(*
 * Simulacion_Trifasico_MPC_v8_M6_it10_opt_S71200.scl
 *
 * Base: Simulacion_Trifasico_MPC_v8_M6_it10_opt_OB100ms_DIAG.scl (PLC Coder 24.1,
 * variante f: Parametros_MPC_v8, M = 6, P = 200, tope de 10 iteraciones, Kr 18x3,
 * divisor desactivado, instrumentacion [DIAG] con RUNTIME).
 *
 * MODIFICADO para S7-1200 (memoria de trabajo). La ley de control no cambia:
 *  1. Kr, Hinv, Ac y Linv pasan a valores iniciales de la declaracion. Se
 *     elimina el bloque need_init, que las cargaba con 2144 asignaciones.
 *  2. rseq pasa de 600 a 3 elementos (solo se usan rseq[0..2]) y se elimina
 *     vseq (201 unos que no se usaban); v sigue valiendo 1.0.
 *  3. Se eliminan las copias QQ y RR: se leen directamente i0_qr.b_Q y i0_qr.b_R.
 *  4. Los arreglos de solo lectura pasan de VAR_INPUT (copia en cada llamada)
 *     a VAR_IN_OUT (referencia): qr.b_A, xgemv.b_A (x se elimina porque en qr
 *     siempre es el mismo arreglo que b_A), mpc_clipping.b_Mlim
 *     y b_Mrows, abs_g.x, b_abs.x, maximum2.x.
 *  5. Bloques con los nombres del proyecto (sufijo _MPC; MPC_3 -> MPC_Control).
 *  v2 (para bajar del 100 % en la CPU 1212C), resultados identicos:
 *  6. Ac separada en AcS (SINT, columnas 0..17, valores -1/0/1) y AcSlack (REAL,
 *     columna 18); cada producto suma la columna 18 al final, en el mismo orden.
 *  7. Se elimina U: en el lazo se usa -b_H (negacion exacta) y en el arranque
 *     en caliente se guarda en TL, que se recalcula antes de volver a leerse.
 *  8. qr factoriza en el sitio sobre RLinv (sin la copia c_A).
 *  9. RLinv, TL y b_D pasan a VAR_TEMP (4332 B de pila local; limite 6 KB).
 * 10. d_a pasa de INT a SINT (valores -1/0/1).
 *  LLAMAR DESDE UN OB CICLICO DE 100 ms. Requiere el DB global Diag_HIL.
 *
 * Model name                      : Simulacion_Trifasico_MPC_v6
 * Model version                   : 1.95
 * Model creator                   : Ivan
 * Model last modified by          : Ivan
 * Model last modified on          : Tue Sep 22 00:34:01 2026
 * Model sample time               : 0.01s
 * Subsystem name                  : Simulacion_Trifasico_MPC_v6/MPC_3
 * Subsystem sample time           : 0.01s
 * Simulink PLC Coder version      : 24.1 (R2024a) 19-Nov-2023
 * ST code generated on            : Tue Sep 22 02:35:18 2026
 *
 * Target IDE selection            : Siemens TIA Portal
 * Test Bench included             : No
 *
 * MODIFICADO (post-proceso), variante f: Parametros_MPC_v8 con M = 6 y tope de 10 iteraciones (P = 200):
 *  - Kr reducida de 18x600 a 18x3: 54 operaciones por ejecucion en lugar de 10800.
 *  - Contador en DB propio: PLCGlobalVarMPC.plc_ts_counter_MPC
 *  - Divisor desactivado: el MPC ejecuta en cada llamada.
 *    LLAMAR DESDE UN OB CICLICO DE 100 ms (100000 us).
 *
 * MODIFICADO: instrumentacion de tiempo con RUNTIME (lineas marcadas [DIAG]).
 *  - Mide el paso completo del MPC: estimador + QP + recorte.
 *  - Registra el estado del QP: iteraciones, llegadas al tope e infactibles.
 *  - Requiere el DB global Diag_HIL (Diag_HIL.scl) en el proyecto.
 *  - La ley de control no cambia.
 *
 *)
DATA_BLOCK PLCGlobalVarMPC
STRUCT
    plc_ts_counter_MPC: DINT;
END_STRUCT
BEGIN
END_DATA_BLOCK
FUNCTION_BLOCK abs_g_MPC
VAR_OUTPUT
    y: ARRAY [0..71] OF REAL;
END_VAR
VAR_IN_OUT
    x: ARRAY [0..71] OF REAL;   (* solo lectura *)
END_VAR
VAR
    k: DINT;
END_VAR
FOR k := 0 TO 71 DO
    y[k] := ABS(x[k]);
END_FOR;
END_FUNCTION_BLOCK
FUNCTION_BLOCK b_abs_MPC
VAR_OUTPUT
    y: ARRAY [0..18] OF REAL;
END_VAR
VAR_IN_OUT
    x: ARRAY [0..18] OF REAL;   (* solo lectura *)
END_VAR
VAR
    k: DINT;
END_VAR
FOR k := 0 TO 18 DO
    y[k] := ABS(x[k]);
END_FOR;
END_FUNCTION_BLOCK
FUNCTION_BLOCK maximum2_MPC
VAR_INPUT
    y: REAL;
END_VAR
VAR_OUTPUT
    ex: ARRAY [0..71] OF REAL;
END_VAR
VAR_IN_OUT
    x: ARRAY [0..71] OF REAL;   (* solo lectura *)
END_VAR
VAR
    k: DINT;
END_VAR
FOR k := 0 TO 71 DO
    ex[k] := MAX(IN1:=x[k], IN2:=y);
END_FOR;
END_FUNCTION_BLOCK
FUNCTION_BLOCK mpc_clipping_MPC
VAR_INPUT
    uk: ARRAY [0..2] OF REAL;
    uk1: ARRAY [0..2] OF REAL;
    b_uoff: ARRAY [0..2] OF REAL;
    b_ny: DINT;
    b_degrees: DINT;
END_VAR
VAR_OUTPUT
    uk_clipped: ARRAY [0..2] OF REAL;
END_VAR
VAR_IN_OUT
    b_Mlim: ARRAY [0..71] OF REAL;   (* solo lectura *)
    b_Mrows: ARRAY [0..71] OF DINT;  (* solo lectura *)
END_VAR
VAR
    nylim: DINT;
    umax: ARRAY [0..2] OF REAL;
    umin: ARRAY [0..2] OF REAL;
    dumin: ARRAY [0..2] OF REAL;
    dumax: ARRAY [0..2] OF REAL;
    iu: DINT;
    du: REAL;
    b_i: DINT;
    tmp: DINT;
    temp1: BOOL;
    temp2: BOOL;
    temp3: BOOL;
END_VAR
nylim := (400 * b_ny) + 1200;
uk_clipped[0] := uk[0];
umax[0] := 3.4028234663852886E+37;
umin[0] := -3.4028234663852886E+37;
dumin[0] := -3.4028234663852886E+37;
dumax[0] := 3.4028234663852886E+37;
uk_clipped[1] := uk[1];
umax[1] := 3.4028234663852886E+37;
umin[1] := -3.4028234663852886E+37;
dumin[1] := -3.4028234663852886E+37;
dumax[1] := 3.4028234663852886E+37;
uk_clipped[2] := uk[2];
umax[2] := 3.4028234663852886E+37;
umin[2] := -3.4028234663852886E+37;
dumin[2] := -3.4028234663852886E+37;
dumax[2] := 3.4028234663852886E+37;
FOR b_i := 0 TO 71 DO
    iu := b_Mrows[b_i];
    temp1 := FALSE;
    temp2 := FALSE;
    temp3 := FALSE;
    IF iu > (nylim - 1200) THEN
        IF iu <= (nylim - 1197) THEN
            iu := (iu - nylim) + 1199;
            umax[iu] := b_Mlim[b_i] + b_uoff[iu];
        ELSE
            temp3 := TRUE;
        END_IF;
    ELSE
        temp3 := TRUE;
    END_IF;
    IF temp3 THEN
        IF iu > (nylim - 600) THEN
            IF iu <= (nylim - 597) THEN
                iu := (iu - nylim) + 599;
                umin[iu] := ( -b_Mlim[b_i]) + b_uoff[iu];
            ELSE
                temp2 := TRUE;
            END_IF;
        ELSE
            temp2 := TRUE;
        END_IF;
    END_IF;
    IF temp2 THEN
        IF iu > nylim THEN
            IF iu <= (nylim + 3) THEN
                dumax[(iu - nylim) - 1] := b_Mlim[b_i];
            ELSE
                temp1 := TRUE;
            END_IF;
        ELSE
            temp1 := TRUE;
        END_IF;
    END_IF;
    IF temp1 THEN
        tmp := nylim + b_degrees;
        IF iu > (tmp - 1) THEN
            IF iu <= (tmp + 2) THEN
                dumin[(iu - nylim) - b_degrees] :=  -b_Mlim[b_i];
            END_IF;
        END_IF;
    END_IF;
END_FOR;
du := uk[0] - uk1[0];
IF du > dumax[0] THEN
    uk_clipped[0] := uk1[0] + dumax[0];
ELSIF du < dumin[0] THEN
    uk_clipped[0] := uk1[0] + dumin[0];
END_IF;
IF uk_clipped[0] > umax[0] THEN
    uk_clipped[0] := umax[0];
ELSIF uk_clipped[0] < umin[0] THEN
    uk_clipped[0] := umin[0];
END_IF;
du := uk[1] - uk1[1];
IF du > dumax[1] THEN
    uk_clipped[1] := uk1[1] + dumax[1];
ELSIF du < dumin[1] THEN
    uk_clipped[1] := uk1[1] + dumin[1];
END_IF;
IF uk_clipped[1] > umax[1] THEN
    uk_clipped[1] := umax[1];
ELSIF uk_clipped[1] < umin[1] THEN
    uk_clipped[1] := umin[1];
END_IF;
du := uk[2] - uk1[2];
IF du > dumax[2] THEN
    uk_clipped[2] := uk1[2] + dumax[2];
ELSIF du < dumin[2] THEN
    uk_clipped[2] := uk1[2] + dumin[2];
END_IF;
IF uk_clipped[2] > umax[2] THEN
    uk_clipped[2] := umax[2];
ELSIF uk_clipped[2] < umin[2] THEN
    uk_clipped[2] := umin[2];
END_IF;
END_FUNCTION_BLOCK
FUNCTION maximum_MPC: REAL
VAR_INPUT
    x: ARRAY [0..18] OF REAL;
END_VAR
VAR_TEMP
    k: DINT;
    x_0: REAL;
END_VAR
maximum_MPC := x[0];
FOR k := 0 TO 17 DO
    x_0 := x[k + 1];
    IF maximum_MPC < x_0 THEN
        maximum_MPC := x_0;
    END_IF;
END_FOR;
END_FUNCTION
FUNCTION_BLOCK DropConstraint_MPC
VAR_INPUT
    kDrop: DINT;
END_VAR
VAR_IN_OUT
    iA: ARRAY [0..71] OF BOOL;
    nA: DINT;
    iC: ARRAY [0..71] OF DINT;
END_VAR
VAR
    b_i: DINT;
END_VAR
IF kDrop > 0 THEN
    iA[iC[kDrop - 1] - 1] := FALSE;
    IF kDrop < nA THEN
        b_i := kDrop;
        WHILE b_i <= (nA - 1) DO
            iC[b_i - 1] := iC[b_i];
            b_i := b_i + 1;
        END_WHILE;
    END_IF;
    iC[nA - 1] := 0;
    nA := nA - 1;
END_IF;
END_FUNCTION_BLOCK
FUNCTION mtimes_MPC: REAL
VAR_INPUT
    b_A: ARRAY [0..18] OF REAL;
    B: ARRAY [0..18] OF REAL;
END_VAR
VAR_TEMP
    k: DINT;
END_VAR
mtimes_MPC := 0.0;
FOR k := 0 TO 18 DO
    mtimes_MPC := (b_A[k] * B[k]) + mtimes_MPC;
END_FOR;
END_FUNCTION
FUNCTION xnrm2_MPC: REAL
VAR_INPUT
    b_n: DINT;
    x: ARRAY [0..360] OF REAL;
    ix0: DINT;
END_VAR
VAR_TEMP
    b_scale: REAL;
    kend: DINT;
    absxk: REAL;
    t: REAL;
    k: DINT;
END_VAR
xnrm2_MPC := 0.0;
IF b_n >= 1 THEN
    IF b_n = 1 THEN
        xnrm2_MPC := ABS(x[ix0 - 1]);
    ELSE
        b_scale := 1.1754943508222875E-37;
        kend := (ix0 + b_n) - 1;
        k := ix0;
        WHILE k <= kend DO
            absxk := ABS(x[k - 1]);
            IF absxk > b_scale THEN
                t := b_scale / absxk;
                xnrm2_MPC := ((xnrm2_MPC * t) * t) + 1.0;
                b_scale := absxk;
            ELSE
                t := absxk / b_scale;
                xnrm2_MPC := (t * t) + xnrm2_MPC;
            END_IF;
            k := k + 1;
        END_WHILE;
        xnrm2_MPC := b_scale * SQRT(xnrm2_MPC);
    END_IF;
END_IF;
END_FUNCTION
FUNCTION_BLOCK xgerc_MPC
VAR_INPUT
    b_m: DINT;
    b_n: DINT;
    alpha1: REAL;
    ix0: DINT;
    y: ARRAY [0..18] OF REAL;
    ia0: DINT;
END_VAR
VAR_IN_OUT
    b_A: ARRAY [0..360] OF REAL;
END_VAR
VAR
    jA: DINT;
    jy: DINT;
    temp: REAL;
    ix: DINT;
    j: DINT;
    b_b: DINT;
    ijA: DINT;
END_VAR
IF alpha1 <> 0.0 THEN
    jA := ia0 - 1;
    jy := 0;
    j := 0;
    WHILE j <= (b_n - 1) DO
        IF y[jy] <> 0.0 THEN
            temp := y[jy] * alpha1;
            ix := ix0;
            ijA := jA;
            b_b := b_m + jA;
            WHILE (ijA + 1) <= b_b DO
                b_A[ijA] := (b_A[ix - 1] * temp) + b_A[ijA];
                ix := ix + 1;
                ijA := ijA + 1;
            END_WHILE;
        END_IF;
        jy := jy + 1;
        jA := jA + 19;
        j := j + 1;
    END_WHILE;
END_IF;
END_FUNCTION_BLOCK
FUNCTION_BLOCK xgemv_MPC
VAR_INPUT
    b_m: DINT;
    b_n: DINT;
    ia0: DINT;
    ix0: DINT;
END_VAR
VAR_IN_OUT
    y: ARRAY [0..18] OF REAL;
    b_A: ARRAY [0..360] OF REAL;   (* solo lectura, por referencia; hace tambien de x: en qr siempre x = b_A = c_A *)
END_VAR
VAR
    ix: DINT;
    b_c: REAL;
    b_iy: DINT;
    b_b: DINT;
    iac: DINT;
    b_d: DINT;
    ia: DINT;
END_VAR
IF (b_m <> 0) AND (b_n <> 0) THEN
    b_iy := 0;
    WHILE b_iy <= (b_n - 1) DO
        y[b_iy] := 0.0;
        b_iy := b_iy + 1;
    END_WHILE;
    b_iy := 0;
    b_b := ((b_n - 1) * 19) + ia0;
    iac := ia0;
    WHILE iac <= b_b DO
        ix := ix0;
        b_c := 0.0;
        b_d := (iac + b_m) - 1;
        ia := iac;
        WHILE ia <= b_d DO
            b_c := (b_A[ia - 1] * b_A[ix - 1]) + b_c;
            ix := ix + 1;
            ia := ia + 1;
        END_WHILE;
        y[b_iy] := y[b_iy] + b_c;
        b_iy := b_iy + 1;
        iac := iac + 19;
    END_WHILE;
END_IF;
END_FUNCTION_BLOCK
FUNCTION_BLOCK qr_MPC
VAR_OUTPUT
    b_Q: ARRAY [0..360] OF REAL;
    b_R: ARRAY [0..360] OF REAL;
END_VAR
VAR_IN_OUT
    b_A: ARRAY [0..360] OF REAL;   (* se factoriza en el sitio: el llamador no vuelve a leer RLinv sin ponerla a cero *)
END_VAR
VAR
    i0_xgemv: xgemv_MPC;
    i0_xgerc: xgerc_MPC;
    tau: ARRAY [0..18] OF REAL;
    itau: DINT;
    work: ARRAY [0..18] OF REAL;
    ii: DINT;
    atmp: REAL;
    beta1: REAL;
    knt: DINT;
    c_lastc: DINT;
    coltop: DINT;
    b_coltop: DINT;
    c_A_0: REAL;
    a: REAL;
    exitg1: DINT;
    exitg2: DINT;
    temp7: REAL;
END_VAR
FOR ii := 0 TO 18 DO
    tau[ii] := 0.0;
    work[ii] := 0.0;
END_FOR;
FOR itau := 0 TO 18 DO
    ii := (itau * 19) + itau;
    IF (itau + 1) < 19 THEN
        atmp := b_A[ii];
        tau[itau] := 0.0;
        beta1 := xnrm2_MPC(b_n := 18 - itau, x := b_A, ix0 := ii + 2);
        IF beta1 <> 0.0 THEN
            c_A_0 := b_A[ii];
            a := ABS(c_A_0);
            beta1 := ABS(beta1);
            IF a < beta1 THEN
                a := a / beta1;
                beta1 := SQRT((a * a) + 1.0) * beta1;
            ELSIF a > beta1 THEN
                beta1 := beta1 / a;
                beta1 := SQRT((beta1 * beta1) + 1.0) * a;
            ELSE
                beta1 := a * 1.4142135623730951;
            END_IF;
            IF c_A_0 >= 0.0 THEN
                beta1 :=  -beta1;
            END_IF;
            IF ABS(beta1) < 1.1754943508222875E-37 THEN
                knt := 0;
                REPEAT
                    exitg1 := 0;
                    knt := knt + 1;
                    c_lastc := (ii - itau) + 19;
                    b_coltop := ii + 1;
                    WHILE (b_coltop + 1) <= c_lastc DO
                        b_A[b_coltop] := 3.4028234663852886E+37 * b_A[b_coltop];
                        b_coltop := b_coltop + 1;
                    END_WHILE;
                    beta1 := beta1 * 3.4028234663852886E+37;
                    atmp := atmp * 3.4028234663852886E+37;
                    IF ABS(beta1) < 1.1754943508222875E-37 THEN
                        IF knt < 20 THEN
                            ;
                            ;
                        ELSE
                            exitg1 := 1;
                        END_IF;
                    ELSE
                        exitg1 := 1;
                    END_IF;
                UNTIL NOT(exitg1 = 0)
                END_REPEAT;
                a := ABS(atmp);
                temp7 := xnrm2_MPC(b_n := 18 - itau, x := b_A, ix0 := ii + 2);
                beta1 := ABS(temp7);
                IF a < beta1 THEN
                    a := a / beta1;
                    beta1 := SQRT((a * a) + 1.0) * beta1;
                ELSIF a > beta1 THEN
                    beta1 := beta1 / a;
                    beta1 := SQRT((beta1 * beta1) + 1.0) * a;
                ELSE
                    beta1 := a * 1.4142135623730951;
                END_IF;
                IF atmp >= 0.0 THEN
                    beta1 :=  -beta1;
                END_IF;
                tau[itau] := (beta1 - atmp) / beta1;
                atmp := 1.0 / (atmp - beta1);
                b_coltop := ii + 1;
                WHILE (b_coltop + 1) <= c_lastc DO
                    b_A[b_coltop] := atmp * b_A[b_coltop];
                    b_coltop := b_coltop + 1;
                END_WHILE;
                c_lastc := 0;
                WHILE c_lastc <= (knt - 1) DO
                    beta1 := beta1 * 1.1754943508222875E-37;
                    c_lastc := c_lastc + 1;
                END_WHILE;
                atmp := beta1;
            ELSE
                tau[itau] := (beta1 - c_A_0) / beta1;
                atmp := 1.0 / (c_A_0 - beta1);
                knt := (ii - itau) + 19;
                c_lastc := ii + 1;
                WHILE (c_lastc + 1) <= knt DO
                    b_A[c_lastc] := atmp * b_A[c_lastc];
                    c_lastc := c_lastc + 1;
                END_WHILE;
                atmp := beta1;
            END_IF;
        END_IF;
        b_A[ii] := 1.0;
        IF tau[itau] <> 0.0 THEN
            knt := 19 - itau;
            c_lastc := (ii - itau) + 18;
            REPEAT
                exitg1 := 0;
                IF knt > 0 THEN
                    IF b_A[c_lastc] = 0.0 THEN
                        knt := knt - 1;
                        c_lastc := c_lastc - 1;
                    ELSE
                        exitg1 := 1;
                    END_IF;
                ELSE
                    exitg1 := 1;
                END_IF;
            UNTIL NOT(exitg1 = 0)
            END_REPEAT;
            c_lastc := 18 - itau;
            REPEAT
                exitg2 := 0;
                IF c_lastc > 0 THEN
                    b_coltop := (((c_lastc - 1) * 19) + ii) + 19;
                    coltop := b_coltop;
                    REPEAT
                        exitg1 := 0;
                        IF (coltop + 1) <= (b_coltop + knt) THEN
                            IF b_A[coltop] <> 0.0 THEN
                                exitg1 := 1;
                            ELSE
                                coltop := coltop + 1;
                            END_IF;
                        ELSE
                            c_lastc := c_lastc - 1;
                            exitg1 := 2;
                        END_IF;
                    UNTIL NOT(exitg1 = 0)
                    END_REPEAT;
                    IF exitg1 = 1 THEN
                        exitg2 := 1;
                    END_IF;
                ELSE
                    exitg2 := 1;
                END_IF;
            UNTIL NOT(exitg2 = 0)
            END_REPEAT;
        ELSE
            knt := 0;
            c_lastc := 0;
        END_IF;
        IF knt > 0 THEN
            i0_xgemv(b_m := knt, b_n := c_lastc, b_A := b_A, ia0 := ii + 20, ix0 := ii + 1, y := work);
            i0_xgerc(b_m := knt, b_n := c_lastc, alpha1 :=  -tau[itau], ix0 := ii + 1, y := work, b_A := b_A, ia0 := ii + 20)
                ;
        END_IF;
        b_A[ii] := atmp;
    ELSE
        tau[18] := 0.0;
    END_IF;
END_FOR;
FOR itau := 0 TO 18 DO
    ii := 0;
    WHILE ii <= itau DO
        b_R[ii + (19 * itau)] := b_A[(19 * itau) + ii];
        ii := ii + 1;
    END_WHILE;
    ii := itau + 1;
    WHILE (ii + 1) < 20 DO
        b_R[ii + (19 * itau)] := 0.0;
        ii := ii + 1;
    END_WHILE;
    work[itau] := 0.0;
END_FOR;
FOR ii := 18 TO 0 BY -1 DO
    knt := ((ii * 19) + ii) + 20;
    IF (ii + 1) < 19 THEN
        b_A[knt - 20] := 1.0;
        IF tau[ii] <> 0.0 THEN
            c_lastc := 19 - ii;
            b_coltop := knt - ii;
            REPEAT
                exitg1 := 0;
                IF c_lastc > 0 THEN
                    IF b_A[b_coltop - 2] = 0.0 THEN
                        c_lastc := c_lastc - 1;
                        b_coltop := b_coltop - 1;
                    ELSE
                        exitg1 := 1;
                    END_IF;
                ELSE
                    exitg1 := 1;
                END_IF;
            UNTIL NOT(exitg1 = 0)
            END_REPEAT;
            b_coltop := 18 - ii;
            REPEAT
                exitg2 := 0;
                IF b_coltop > 0 THEN
                    coltop := ((b_coltop - 1) * 19) + knt;
                    itau := coltop;
                    REPEAT
                        exitg1 := 0;
                        IF itau <= ((coltop + c_lastc) - 1) THEN
                            IF b_A[itau - 1] <> 0.0 THEN
                                exitg1 := 1;
                            ELSE
                                itau := itau + 1;
                            END_IF;
                        ELSE
                            b_coltop := b_coltop - 1;
                            exitg1 := 2;
                        END_IF;
                    UNTIL NOT(exitg1 = 0)
                    END_REPEAT;
                    IF exitg1 = 1 THEN
                        exitg2 := 1;
                    END_IF;
                ELSE
                    exitg2 := 1;
                END_IF;
            UNTIL NOT(exitg2 = 0)
            END_REPEAT;
        ELSE
            c_lastc := 0;
            b_coltop := 0;
        END_IF;
        IF c_lastc > 0 THEN
            i0_xgemv(b_m := c_lastc, b_n := b_coltop, b_A := b_A, ia0 := knt, ix0 := knt - 19, y := work);
            i0_xgerc(b_m := c_lastc, b_n := b_coltop, alpha1 :=  -tau[ii], ix0 := knt - 19, y := work, b_A := b_A, ia0 := knt)
                ;
        END_IF;
        c_lastc := (knt - ii) - 1;
        b_coltop := knt - 19;
        WHILE (b_coltop + 1) <= c_lastc DO
            b_A[b_coltop] := ( -tau[ii]) * b_A[b_coltop];
            b_coltop := b_coltop + 1;
        END_WHILE;
    END_IF;
    b_A[knt - 20] := 1.0 - tau[ii];
    c_lastc := 0;
    WHILE c_lastc <= (ii - 1) DO
        b_A[(knt - c_lastc) - 21] := 0.0;
        c_lastc := c_lastc + 1;
    END_WHILE;
END_FOR;
FOR ii := 0 TO 360 DO
    b_Q[ii] := b_A[ii];
END_FOR;
END_FUNCTION_BLOCK
FUNCTION b_norm_MPC: REAL
VAR_INPUT
    x: ARRAY [0..18] OF REAL;
END_VAR
VAR_TEMP
    b_scale: REAL;
    absxk: REAL;
    t: REAL;
    k: DINT;
END_VAR
b_norm_MPC := 0.0;
b_scale := 1.1754943508222875E-37;
FOR k := 0 TO 18 DO
    absxk := ABS(x[k]);
    IF absxk > b_scale THEN
        t := b_scale / absxk;
        b_norm_MPC := ((b_norm_MPC * t) * t) + 1.0;
        b_scale := absxk;
    ELSE
        t := absxk / b_scale;
        b_norm_MPC := (t * t) + b_norm_MPC;
    END_IF;
END_FOR;
b_norm_MPC := b_scale * SQRT(b_norm_MPC);
END_FUNCTION
FUNCTION_BLOCK mpcblock_refmd_MPC
VAR_INPUT
    b_ref: ARRAY [0..2] OF REAL;
    b_yoff: ARRAY [0..2] OF REAL;
    b_RYscale: ARRAY [0..2] OF REAL;
END_VAR
VAR_OUTPUT
    rseq: ARRAY [0..2] OF REAL;   (* antes 0..599: solo se usan rseq[0..2] *)
    v: REAL;
END_VAR
VAR
    b_i: DINT;
    ref_0: REAL;
    ref_1: REAL;
    ref_2: REAL;
    b_RYscale_0: REAL;
    b_RYscale_1: REAL;
    b_RYscale_2: REAL;
    b_yoff_0: REAL;
    b_yoff_1: REAL;
    b_yoff_2: REAL;
END_VAR
ref_0 := b_ref[0];
ref_1 := b_ref[1];
ref_2 := b_ref[2];
b_RYscale_0 := b_RYscale[0];
b_RYscale_1 := b_RYscale[1];
b_RYscale_2 := b_RYscale[2];
b_yoff_0 := b_yoff[0];
b_yoff_1 := b_yoff[1];
b_yoff_2 := b_yoff[2];
FOR b_i := 0 TO 0 DO    (* solo rseq[0..2] se usa *)
    rseq[b_i * 3] := (ref_0 * b_RYscale_0) - b_yoff_0;
    rseq[(b_i * 3) + 1] := (ref_1 * b_RYscale_1) - b_yoff_1;
    rseq[(b_i * 3) + 2] := (ref_2 * b_RYscale_2) - b_yoff_2;
END_FOR;
v := 1.0;
END_FUNCTION_BLOCK
FUNCTION rt_floord_MPC: REAL
VAR_INPUT
    u: REAL;
END_VAR
rt_floord_MPC := DINT_TO_REAL(TRUNC(u));
IF u = rt_floord_MPC THEN
    rt_floord_MPC := u;
ELSIF u < 0.0 THEN
    rt_floord_MPC := rt_floord_MPC - 1.0;
END_IF;
END_FUNCTION
FUNCTION_BLOCK MPC_Control
VAR_INPUT
    ssMethodType: INT;
    moorx: ARRAY [0..2] OF REAL;
    b_ref: ARRAY [0..2] OF REAL;
END_VAR
VAR_OUTPUT
    mv: ARRAY [0..2] OF REAL;
END_VAR
VAR
    Memory_PreviousInput: ARRAY [0..71] OF BOOL;
    last_x_PreviousInput: ARRAY [0..6] OF REAL;
    last_mv_DSTATE: ARRAY [0..2] OF REAL;
    MathFunction: ARRAY [0..2] OF REAL;
    MathFunction1: ARRAY [0..2] OF REAL;
    MathFunction2: ARRAY [0..2] OF REAL;
    c_last_x_InitialCond: ARRAY [0..6] OF REAL := [0.47374550049727165,0.8,0.72,255106.009,0.0,0.0,0.0];
    MPC_3_b_myoff: ARRAY [0..2] OF REAL := [0.8,0.72,3.7];
    MPC_3_b_RYscale: ARRAY [0..2] OF REAL := [1.0,1.0,0.1];
    MPC_3_b_xoff: ARRAY [0..6] OF REAL := [0.47374550049727165,0.8,0.72,255106.009,0.0,0.0,0.0];
    b_a: ARRAY [0..20] OF REAL := [0.0,0.0,0.0,1.0,0.0,0.0,0.0,1.0,0.0,0.0,0.0,1.4503774389728313E-5,0.0,0.0,0.0,0.0,0.0,0.0,0.0,
        0.0,0.0];
    MPC_3_c_a: ARRAY [0..20] OF REAL := [-0.0772292027423523,0.12077646327456022,0.0038948707411090538,1352.9330397447068,
        3.4881337436777948,-1.3447885799979777,-1.1731438171327024,0.269035613232814,0.0038948707411099914,0.09786695730401461,
        348.05070726193321,0.11111867957141662,2.7949959088743932,-2.8155753844244291,0.059593437249509731,0.01962263557286395,
        0.0050480489343075492,14331.413461436903,1.6106730948140586,2.3311020292522353,2.408935193579286];
    d_a: ARRAY [0..215] OF SINT := [-1,0,0,-1,0,0,-1,0,0,-1,0,0,-1,0,0,-1,0,0,1,0,0,1,0,0,1,0,0,1,0,0,1,0,0,1,0,0,0,0,0,0,0,0,0,0,0,
        0,0,0,0,0,0,0,0,0,0,0,0,0,0,0,0,0,0,0,0,0,0,0,0,0,0,0,0,-1,0,0,-1,0,0,-1,0,0,-1,0,0,-1,0,0,-1,0,0,1,0,0,1,0,0,1,0,0,
        1,0,0,1,0,0,1,0,0,0,0,0,0,0,0,0,0,0,0,0,0,0,0,0,0,0,0,0,0,0,0,0,0,0,0,0,0,0,0,0,0,0,0,0,0,0,-1,0,0,-1,0,0,-1,0,0,-1,
        0,0,-1,0,0,-1,0,0,1,0,0,1,0,0,1,0,0,1,0,0,1,0,0,1,0,0,0,0,0,0,0,0,0,0,0,0,0,0,0,0,0,0,0,0,0,0,0,0,0,0,0,0,0,0,0,0,0,
        0,0,0];
    MPC_3_b_Mlim: ARRAY [0..71] OF REAL := [0.333871875208127,0.752014397384409,0.515635973890735,0.333871875208127,
        0.752014397384409,0.515635973890735,0.333871875208127,0.752014397384409,0.515635973890735,0.333871875208127,0.752014397384409,
        0.515635973890735,0.333871875208127,0.752014397384409,0.515635973890735,0.333871875208127,0.752014397384409,0.515635973890735,
        0.636128124791873,0.21798560261559102,0.45436402610926496,0.636128124791873,0.21798560261559102,0.45436402610926496,
        0.636128124791873,0.21798560261559102,0.45436402610926496,0.636128124791873,0.21798560261559102,0.45436402610926496,
        0.636128124791873,0.21798560261559102,0.45436402610926496,0.636128124791873,0.21798560261559102,0.45436402610926496,0.035,0.015,
        0.03,0.035,0.015,0.03,0.035,0.015,0.03,0.035,0.015,0.03,0.035,0.015,0.03,0.035,0.015,0.03,0.035,0.015,0.03,0.035,0.015,
        0.03,0.035,0.015,0.03,0.035,0.015,0.03,0.035,0.015,0.03,0.035,0.015,0.03];
    MPC_3_b_Kx: ARRAY [0..125] OF REAL := [-7716.2321024491939,-10901.008671532656,-4264.9443651421188,0.001588040838629834,
        -2543.7442519006345,-1928.3474040587275,19.549174933816971,-44534.108859815329,-44494.776516572136,-26655.405567238093,
        0.0095121063518449449,-8398.6455416316712,-10368.267059564856,158.86185382546796,877.70571831208667,990.07022975809957,
        474.28108255756024,-0.0035701887162486057,96.5496604150103,99.981804413078876,-126.88330315000997,-7621.9188571763643,
        -10775.120625744157,-4206.5654308225376,0.0015700336455973293,-2519.1535379237243,-1907.0052261791157,19.280661326360363,
        -44188.119848216615,-44149.311125111242,-26390.969999054745,0.0094459267062587185,-8342.2703225681144,-10298.597291206755,
        157.85188650166057,864.95022738088733,975.66168439016542,466.81791298662728,-0.0035336819710021609,94.4868041100247,
        97.85316386731445,-125.93879584019494,-7528.1481322542822,-10649.931335099882,-4148.6767278274638,0.0015521046865827432,
        -2494.6400124657093,-1885.7587961853874,19.013959064141872,-43842.116288935795,-43803.826542255309,-26127.843886728973,
        0.0093796925467878947,-8285.8873550992248,-10228.919297363989,156.8419334382582,852.3095979437818,961.384106890396,459.43616436780036,
        -0.003497369852713806,92.447632839384539,95.74911914998566,-124.99418234183436,-7434.9230075303494,-10525.443894660129,
        -4091.2769580451954,0.0015342547665065048,-2470.2045128943837,-1864.6086925692725,18.749068146716176,-43496.122480806749,
        -43458.347088410825,-25866.027371158609,0.0093134067140901722,-8229.4967444644935,-10159.23320514503,155.83198146211291,
        839.78359704931961,947.23718912342133,452.13534732790527,-0.0034612522993006938,90.432068275420264,93.669582511506164,
        -124.04951211934259,-7342.2465048437853,-10401.661341488485,-4034.3648155478659,0.0015164846849855819,-2445.8478788030538,
        -1843.5554965261258,18.485988665509439,-43150.162591337648,-43112.896952629555,-25605.520593125708,0.0092470720701684772,
        -8173.0986508239621,-10089.539209226115,154.82201815145478,827.37198501561852,933.22061617028339,444.91497290855955,
        -0.0034253292477243787,88.440031602080353,91.614465843510473,-123.10483463065196,-7250.1215881048793,-10278.586654731167,
        -3977.9389865477651,0.00149879523623798,-2421.5709518529893,-1822.5997917608677,18.224720801734843,-42804.2606574284,
        -42767.500193326021,-25346.323693295184,0.0091806914982297729,-8116.6932889508143,-10019.83757147498,153.81203184149854,
        815.07451548496078,919.33406638300414,437.7745525706747,-0.0033896006339887937,86.47144350229388,89.5836806634611,
        -122.16019932703135];
    MPC_3_b_Ku1: ARRAY [0..53] OF REAL := [532.9519035819452,1758.7630386838541,-20.218495148255496,1758.7630386838541,
        9920.4082612993716,-164.30092992093171,-20.218495148255496,-164.30092992093171,131.49311423922407,527.80102628666316,
        1737.934860701725,-19.940788232849528,1746.9574860985949,9846.5918503106168,-163.25638356511735,-19.786511752201875,
        -161.71101778484783,130.514941055735,522.666313063715,1717.21838942958,-19.664954679108821,1735.1503109173054,9772.77075083077,
        -162.21185195795246,-19.359488246736596,-159.14605147852319,129.53665804804106,517.54793926655793,1696.6142696551719,
        -19.390994486572826,1723.3415351782228,9698.9487212665517,-161.16732147527,-18.93740822923742,-156.60596908182839,128.55831637410802,
        512.44608071469349,1676.1231380934234,-19.118907749797927,1711.5311924205112,9625.129520129678,-160.12277927000616,
        -18.520255194809877,-154.09070753671722,127.57996718519767,507.36091366067569,1655.7456233405144,-18.848694656201634,
        1699.7193276198914,9551.3169060341625,-159.07821327799945,-18.108012533640888,-151.60020265098143,126.60166162568011];
    MPC_3_b_Kr: ARRAY [0..53] OF REAL := [3186.8373350513389,4275.3677914960599,51.13509990647421,-32.452540397628589,26714.198696645544,72.918687149547608,
        -112.44555961175674,-475.25673471668864,252.72878690712173,3155.2425613858004,4216.8654170260106,50.638144210838703,
        -31.975100691061328,26449.325655557303,72.210143687081711,-110.79080635121332,-467.77820186026861,250.27164490947899,
        3123.8040857581582,4158.8539359264387,50.143499486122451,-31.502311016836352,26185.762042540995,71.504893608304656,
        -109.15217877028672,-460.38123779321489,247.82594499281888,3092.5219240585361,4101.3320539069082,49.651167400702548,
        -31.034149716397167,25923.508020768073,70.802939302930895,-107.52960162200367,-453.06535277614643,245.39169524300604,
        3061.396092190324,4044.2984688129827,49.161149624113243,-30.57059511536292,25662.563753294817,70.104283162373875,
        -105.92299960583885,-445.83005747772961,242.96890375165114,3030.4266060701984,3987.7518705822636,48.673447827046601,
        -30.111625523516803,25402.929403061011,69.408927579747242,-104.33229736767574,-438.67486297920362,240.55757861611488];   (* Kr reducida 18x3 *)
    MPC_3_b_Hinv: ARRAY [0..360] OF REAL := [0.1702344980572631,-0.000316051953237396,-0.0001214533827540456,-0.036345548841276047,-0.00022994447282000675,
        -7.8535204077971989E-5,-0.035434727013087031,-0.00014382977097906262,-3.4945956300716842E-5,-0.034542309014010772,
        -5.7720706811642746E-5,8.813456011776322E-6,-0.03366968301464044,2.8361008307101794E-5,5.2380161360600679E-5,
        -0.032817675154182616,0.00011438593593406882,9.552481608298865E-5,0.0,-0.000316051953237396,0.010547207252793461,
        2.1132487152157335E-5,-0.0001808791608454948,-0.0023314158969080174,1.0330320315621911E-5,-4.9534035220164727E-5,
        -0.0022413766833578007,1.2191170747377299E-7,7.8036147649309862E-5,-0.0021522792952646508,-9.54953740575078E-6,
        0.00020190252942289518,-0.0020644122541486152,-1.8729858790232883E-5,0.0003221473455128597,-0.0019779594821308214,
        -2.7454115420488076E-5,0.0,-0.0001214533827540456,2.1132487152157335E-5,0.30304411821884769,-6.514990994147179E-5,
        2.1728353827661485E-5,-0.064405415788092474,-8.97885060327611E-6,2.2273463510311548E-5,-0.062989706993492336,
        4.65603793551569E-5,2.2723267969727878E-5,-0.061614542822731315,0.00010110834451599296,2.3046591530932414E-5,
        -0.060282635561179215,0.00015444098334013595,2.322473034505095E-5,-0.058995530723217567,0.0,-0.036345548841276047,
        -0.0001808791608454948,-6.514990994147179E-5,0.17176291685304779,-0.00013612744730930092,-4.4560767159202152E-5,
        -0.0350971665966896,-9.13556293645426E-5,-2.2988766629637194E-5,-0.034463114486899891,-4.65576358502461E-5,
        -9.4991020623304764E-7,-0.033843716347050953,-1.7392388529733022E-6,2.1176229123452892E-5,-0.033239892629933931,
        4.3085064069324768E-5,4.3143636253156359E-5,0.0,-0.00022994447282000675,-0.0023314158969080174,2.1728353827661485E-5,
        -0.00013612744730930092,0.010698246530635966,1.2340538427932472E-5,-4.4760194642908621E-5,-0.0022102015392433554,
        3.4084100679808667E-6,4.4173612422238355E-5,-0.00214976861316072,-5.120830508461208E-6,0.00013070925637258645,
        -0.0020899593246978244,-1.3289405671251868E-5,0.00021489433364024608,-0.0020309671075964997,-2.1128873179308238E-5,
        0.0,-7.8535204077971989E-5,1.0330320315621911E-5,-0.064405415788092474,-4.4560767159202152E-5,1.2340538427932472E-5,
        0.3054148208775625,-1.015071319787011E-5,1.4368446176665112E-5,-0.062417276373171432,2.4179024444158472E-5,
        1.636636500723434E-5,-0.061380921474166857,5.8051555293553663E-5,1.8300251292219083E-5,-0.0603809302382588,
        9.1225498596546247E-5,2.0148793762691288E-5,-0.0594190724227041,0.0,-0.035434727013087031,-4.9534035220164727E-5,
        -8.97885060327611E-6,-0.0350971665966896,-4.4760194642908621E-5,-1.015071319787011E-5,0.17273845134311319,
        -3.9976889795088581E-5,-1.0826124612172019E-5,-0.034391366089294419,-3.5166046909618539E-5,-1.0727884762180431E-5,
        -0.0340234548514619,-3.0316948364924829E-5,-1.0252653775071641E-5,-0.033666135978688227,-2.5428615172775216E-5,
        -9.6634672683266118E-6,0.0,-0.00014382977097906262,-0.0022413766833578007,2.2273463510311548E-5,-9.13556293645426E-5,
        -0.0022102015392433554,1.4368446176665112E-5,-3.9976889795088581E-5,0.010790253977071384,6.7106504165377462E-6,
        1.0310200452023578E-5,-0.002147190141859824,-6.7830888060647946E-7,5.9505058354541645E-5,-0.0021154443640503916,
        -7.8370437343924534E-6,0.00010762063469870516,-0.0020839183592772296,-1.4793606326937087E-5,0.0,
        -3.4945956300716842E-5,1.2191170747377299E-7,-0.062989706993492336,-2.2988766629637194E-5,3.4084100679808667E-6,
        -0.062417276373171432,-1.0826124612172019E-5,6.7106504165377462E-6,0.30702802540700186,1.820897001919164E-6,
        1.005184108764361E-5,-0.061176025329871223,1.4557473121748288E-5,1.3395015801887418E-5,-0.060507679924504308,
        2.7124492071147717E-5,1.6716205009836463E-5,-0.059870813633310996,0.0,-0.034542309014010772,7.8036147649309862E-5,
        4.65603793551569E-5,-0.034463114486899891,4.4173612422238355E-5,2.4179024444158472E-5,-0.034391366089294419,
        1.0310200452023578E-5,1.820897001919164E-6,0.17318140332130527,-2.3547509119607678E-5,-2.0255119613621428E-5,
        -0.03420782335043554,-5.7379181065111574E-5,-4.1654408632959635E-5,-0.034095412692558565,-9.1167816691611789E-5,
        -6.2657366574418234E-5,0.0,-5.7720706811642746E-5,-0.0021522792952646508,2.2723267969727878E-5,-4.65576358502461E-5,
        -0.00214976861316072,1.636636500723434E-5,-3.5166046909618539E-5,-0.002147190141859824,1.005184108764361E-5,
        -2.3547509119607678E-5,0.010824871877124352,3.8016754445631412E-6,-1.1714654534696886E-5,-0.0021406660168113629,
        -2.3487140810286621E-6,3.1080884145891323E-7,-0.0021366194369659398,-8.4238697344242429E-6,0.0,8.813456011776322E-6,
        -9.54953740575078E-6,-0.061614542822731315,-9.4991020623304764E-7,-5.120830508461208E-6,-0.061380921474166857,
        -1.0727884762180431E-5,-6.7830888060647946E-7,-0.061176025329871223,-2.0255119613621428E-5,3.8016754445631412E-6,
        0.30790449828673894,-2.9132918265929341E-5,8.3532488641258142E-6,-0.060660620175687734,-3.7638527243085177E-5,
        1.2949735033266653E-5,-0.060348692971084965,0.0,-0.03366968301464044,0.00020190252942289518,0.00010110834451599296,
        -0.033843716347050953,0.00013070925637258645,5.8051555293553663E-5,-0.0340234548514619,5.9505058354541645E-5,
        1.4557473121748288E-5,-0.03420782335043554,-1.1714654534696886E-5,-2.9132918265929341E-5,0.17311211771562424,
        -8.2943372514784056E-5,-7.26451760390996E-5,-0.034526178406331057,-0.00015415495715396418,-0.00011546864934107219,0.0,
        2.8361008307101794E-5,-0.0020644122541486152,2.3046591530932414E-5,-1.7392388529733022E-6,-0.0020899593246978244,
        1.8300251292219083E-5,-3.0316948364924829E-5,-0.0021154443640503916,1.3395015801887418E-5,-5.7379181065111574E-5,
        -0.0021406660168113629,8.3532488641258142E-6,-8.2943372514784056E-5,0.010803886559746703,3.2103542526533054E-6,
        -0.00010704208143625654,-0.0021887753347569921,-1.9842771425297006E-6,0.0,5.2380161360600679E-5,
        -1.8729858790232883E-5,-0.060282635561179215,2.1176229123452892E-5,-1.3289405671251868E-5,-0.0603809302382588,
        -1.0252653775071641E-5,-7.8370437343924534E-6,-0.060507679924504308,-4.1654408632959635E-5,-2.3487140810286621E-6,
        -0.060660620175687734,-7.26451760390996E-5,3.2103542526533054E-6,0.308065547905881,-0.00010270880655031663,
        8.8847998121922669E-6,-0.0608495071191091,0.0,-0.032817675154182616,0.0003221473455128597,0.00015444098334013595,
        -0.033239892629933931,0.00021489433364024608,9.1225498596546247E-5,-0.033666135978688227,0.00010762063469870516,
        2.7124492071147717E-5,-0.034095412692558565,3.1080884145891323E-7,-3.7638527243085177E-5,-0.034526178406331057,
        -0.00010704208143625654,-0.00010270880655031663,0.17255097784265849,-0.00021442620951791223,-0.00016759605920454502,
        0.0,0.00011438593593406882,-0.0019779594821308214,2.322473034505095E-5,4.3085064069324768E-5,-0.0020309671075964997,
        2.0148793762691288E-5,-2.5428615172775216E-5,-0.0020839183592772296,1.6716205009836463E-5,-9.1167816691611789E-5,
        -0.0021366194369659398,1.2949735033266653E-5,-0.00015415495715396418,-0.0021887753347569921,8.8847998121922669E-6,
        -0.00021442620951791223,0.010729219465504205,4.5706825441767981E-6,0.0,9.552481608298865E-5,-2.7454115420488076E-5,
        -0.058995530723217567,4.3143636253156359E-5,-2.1128873179308238E-5,-0.0594190724227041,-9.6634672683266118E-6,
        -1.4793606326937087E-5,-0.059870813633310996,-6.2657366574418234E-5,-8.4238697344242429E-6,-0.060348692971084965,
        -0.00011546864934107219,-1.9842771425297006E-6,-0.0608495071191091,-0.00016759605920454502,4.5706825441767981E-6,
        0.30753298042695221,0.0,0.0,0.0,0.0,0.0,0.0,0.0,0.0,0.0,0.0,0.0,0.0,0.0,0.0,0.0,0.0,0.0,0.0,0.0,
        9.9999999999999974E-6];
    (* Ac (72 x 19, por columnas) separada: columnas 0..17 solo valen -1, 0 o 1 *)
    AcS: ARRAY [0..1295] OF SINT := [-1,0,0,-1,0,0,-1,0,0,-1,0,0,-1,0,0,-1,0,0,1,0,0,1,0,0,1,0,0,1,0,0,1,0,0,1,0,0,-1,0,0,0,0,0,0,0,0,0,0,0,0,0,0,0,0,0,1,
        0,0,0,0,0,0,0,0,0,0,0,0,0,0,0,0,0,0,-1,0,0,-1,0,0,-1,0,0,-1,0,0,-1,0,0,-1,0,0,1,0,0,1,0,0,1,0,0,1,0,0,1,0,0,1,0,0,-1,
        0,0,0,0,0,0,0,0,0,0,0,0,0,0,0,0,0,1,0,0,0,0,0,0,0,0,0,0,0,0,0,0,0,0,0,0,-1,0,0,-1,0,0,-1,0,0,-1,0,0,-1,0,0,-1,0,0,1,0,
        0,1,0,0,1,0,0,1,0,0,1,0,0,1,0,0,-1,0,0,0,0,0,0,0,0,0,0,0,0,0,0,0,0,0,1,0,0,0,0,0,0,0,0,0,0,0,0,0,0,0,0,0,0,-1,0,0,-1,
        0,0,-1,0,0,-1,0,0,-1,0,0,0,0,0,1,0,0,1,0,0,1,0,0,1,0,0,1,0,0,0,0,0,-1,0,0,0,0,0,0,0,0,0,0,0,0,0,0,0,0,0,1,0,0,0,0,0,0,
        0,0,0,0,0,0,0,0,0,0,0,0,-1,0,0,-1,0,0,-1,0,0,-1,0,0,-1,0,0,0,0,0,1,0,0,1,0,0,1,0,0,1,0,0,1,0,0,0,0,0,-1,0,0,0,0,0,0,0,
        0,0,0,0,0,0,0,0,0,0,1,0,0,0,0,0,0,0,0,0,0,0,0,0,0,0,0,0,0,-1,0,0,-1,0,0,-1,0,0,-1,0,0,-1,0,0,0,0,0,1,0,0,1,0,0,1,0,0,
        1,0,0,1,0,0,0,0,0,-1,0,0,0,0,0,0,0,0,0,0,0,0,0,0,0,0,0,1,0,0,0,0,0,0,0,0,0,0,0,0,0,0,0,0,0,0,-1,0,0,-1,0,0,-1,0,0,-1,
        0,0,0,0,0,0,0,0,1,0,0,1,0,0,1,0,0,1,0,0,0,0,0,0,0,0,-1,0,0,0,0,0,0,0,0,0,0,0,0,0,0,0,0,0,1,0,0,0,0,0,0,0,0,0,0,0,0,0,
        0,0,0,0,0,-1,0,0,-1,0,0,-1,0,0,-1,0,0,0,0,0,0,0,0,1,0,0,1,0,0,1,0,0,1,0,0,0,0,0,0,0,0,-1,0,0,0,0,0,0,0,0,0,0,0,0,0,0,
        0,0,0,1,0,0,0,0,0,0,0,0,0,0,0,0,0,0,0,0,0,0,-1,0,0,-1,0,0,-1,0,0,-1,0,0,0,0,0,0,0,0,1,0,0,1,0,0,1,0,0,1,0,0,0,0,0,0,0,
        0,-1,0,0,0,0,0,0,0,0,0,0,0,0,0,0,0,0,0,1,0,0,0,0,0,0,0,0,0,0,0,0,0,0,0,0,0,0,-1,0,0,-1,0,0,-1,0,0,0,0,0,0,0,0,0,0,0,1,
        0,0,1,0,0,1,0,0,0,0,0,0,0,0,0,0,0,-1,0,0,0,0,0,0,0,0,0,0,0,0,0,0,0,0,0,1,0,0,0,0,0,0,0,0,0,0,0,0,0,0,0,0,0,0,-1,0,0,
        -1,0,0,-1,0,0,0,0,0,0,0,0,0,0,0,1,0,0,1,0,0,1,0,0,0,0,0,0,0,0,0,0,0,-1,0,0,0,0,0,0,0,0,0,0,0,0,0,0,0,0,0,1,0,0,0,0,0,
        0,0,0,0,0,0,0,0,0,0,0,0,0,-1,0,0,-1,0,0,-1,0,0,0,0,0,0,0,0,0,0,0,1,0,0,1,0,0,1,0,0,0,0,0,0,0,0,0,0,0,-1,0,0,0,0,0,0,0,
        0,0,0,0,0,0,0,0,0,0,1,0,0,0,0,0,0,0,0,0,0,0,0,0,0,0,0,0,0,-1,0,0,-1,0,0,0,0,0,0,0,0,0,0,0,0,0,0,1,0,0,1,0,0,0,0,0,0,0,
        0,0,0,0,0,0,0,-1,0,0,0,0,0,0,0,0,0,0,0,0,0,0,0,0,0,1,0,0,0,0,0,0,0,0,0,0,0,0,0,0,0,0,0,0,-1,0,0,-1,0,0,0,0,0,0,0,0,0,
        0,0,0,0,0,1,0,0,1,0,0,0,0,0,0,0,0,0,0,0,0,0,0,-1,0,0,0,0,0,0,0,0,0,0,0,0,0,0,0,0,0,1,0,0,0,0,0,0,0,0,0,0,0,0,0,0,0,0,
        0,0,-1,0,0,-1,0,0,0,0,0,0,0,0,0,0,0,0,0,0,1,0,0,1,0,0,0,0,0,0,0,0,0,0,0,0,0,0,-1,0,0,0,0,0,0,0,0,0,0,0,0,0,0,0,0,0,1,
        0,0,0,0,0,0,0,0,0,0,0,0,0,0,0,0,0,0,-1,0,0,0,0,0,0,0,0,0,0,0,0,0,0,0,0,0,1,0,0,0,0,0,0,0,0,0,0,0,0,0,0,0,0,0,-1,0,0,0,
        0,0,0,0,0,0,0,0,0,0,0,0,0,0,1,0,0,0,0,0,0,0,0,0,0,0,0,0,0,0,0,0,0,-1,0,0,0,0,0,0,0,0,0,0,0,0,0,0,0,0,0,1,0,0,0,0,0,0,
        0,0,0,0,0,0,0,0,0,0,0,-1,0,0,0,0,0,0,0,0,0,0,0,0,0,0,0,0,0,1,0,0,0,0,0,0,0,0,0,0,0,0,0,0,0,0,0,0,-1,0,0,0,0,0,0,0,0,0,
        0,0,0,0,0,0,0,0,1,0,0,0,0,0,0,0,0,0,0,0,0,0,0,0,0,0,-1,0,0,0,0,0,0,0,0,0,0,0,0,0,0,0,0,0,1];
    AcSlack: ARRAY [0..71] OF REAL := [0.1,0.1,0.1,0.1,0.1,0.1,0.1,0.1,0.1,0.1,0.1,0.1,0.1,0.1,0.1,0.1,0.1,0.1,0.1,0.1,0.1,0.1,0.1,0.1,0.1,0.1,0.1,0.1,0.1,
        0.1,0.1,0.1,0.1,0.1,0.1,0.1,0.0,0.0,0.0,0.0,0.0,0.0,0.0,0.0,0.0,0.0,0.0,0.0,0.0,0.0,0.0,0.0,0.0,0.0,0.0,0.0,0.0,0.0,
        0.0,0.0,0.0,0.0,0.0,0.0,0.0,0.0,0.0,0.0,0.0,0.0,0.0,0.0];   (* columna 18: holgura *)
    MPC_3_b_uoff: ARRAY [0..2] OF REAL := [0.656128124791873,0.237985602615591,0.474364026109265];
    MPC_3_b_Mrows: ARRAY [0..71] OF DINT := [1201,1202,1203,1204,1205,1206,1207,1208,1209,1210,1211,1212,1213,1214,1215,1216,1217,
        1218,1801,1802,1803,1804,1805,1806,1807,1808,1809,1810,1811,1812,1813,1814,1815,1816,1817,1818,2401,2402,2403,2404,
        2405,2406,2407,2408,2409,2410,2411,2412,2413,2414,2415,2416,2417,2418,2419,2420,2421,2422,2423,2424,2425,2426,2427,
        2428,2429,2430,2431,2432,2433,2434,2435,2436];
    MPC_3_b_Linv: ARRAY [0..360] OF REAL := [0.043122239395521268,-0.05019306519247696,-0.0033206696132972837,-0.31577942830214772,-0.0031471197006212965,
        -0.00020705051348992359,-0.18308150772189805,-0.0014696017526715675,-7.5450474722372636E-5,-0.12889586192277314,
        -0.00059021717051271558,3.8407404253082784E-6,-0.09869296350827321,0.0002261820630442589,8.3395085100205E-5,
        -0.078999376861682777,0.0011042900946144102,0.00017225441484848154,0.0,0.0,0.015347363356332721,0.0020190838633724136,
        -0.00091102072052030891,-0.07901358568341027,6.7218935720810737E-5,-9.1246872819404E-6,-0.045684177963437142,
        -3.9801617956080181E-6,0.00027433939577582988,-0.031987683695103353,-2.7972250421381947E-5,0.00047973300959174817,
        -0.024247405963223941,-4.0683462098209086E-5,0.0006803357457738446,-0.01909559690027262,-4.9506429646829944E-5,0.0,
        0.0,0.0,0.087312641366686636,-0.00043386070373357613,0.001238779140346204,-0.42107641020149239,-6.1807887311560788E-5,
        0.00051363050814862469,-0.24423350048424408,7.3761326011918756E-5,0.00035445285917561705,-0.17220651542065402,
        0.00018273894349911022,0.00028329895418285477,-0.13225134353194426,0.00029556006650442523,0.00023268095887176668,
        -0.10638325243751168,0.0,0.0,0.0,0.0,0.32476352152728083,-0.0022032755395640763,-0.00021807552222073261,
        -0.1826323676701698,-0.0012233193115584247,-0.00011214950035355466,-0.12907314160690159,-0.00073675201931614072,
        -5.3944104655688172E-5,-0.0993319703512495,-0.00021614122189525552,6.5016994885151178E-6,-0.080019318890644078,
        0.00041594529543757932,7.77984415145777E-5,0.0,0.0,0.0,0.0,0.0,0.081196332633548682,9.4178408876197282E-5,
        -0.00018552342484247817,-0.045616373263034124,1.3382645905252523E-5,7.3265273574636073E-5,-0.032161700136474826,
        -1.4106521576734893E-5,0.00024883046634005361,-0.024605618012537182,-2.8451514186729147E-5,0.00041959371575441944,
        -0.019607343607742585,-3.810048357222283E-5,0.0,0.0,0.0,0.0,0.0,0.0,0.43311489522212737,-0.00017825206901915394,
        0.00037846148477057873,-0.24327007517811419,-5.0314671809548014E-5,0.00026963086606063725,-0.17200596953896155,
        4.5079990938181534E-5,0.0002299643325305634,-0.13258611861207259,0.00014267226685941574,0.00020304604787921979,
        -0.10714700086017916,0.0,0.0,0.0,0.0,0.0,0.0,0.0,0.37344065756375838,-0.00097294854471077308,-0.00014891231274351814,
        -0.12927510944801096,-0.00087014142142283494,-0.00011208292497242445,-0.099986751616224556,-0.00063795107819119646,
        -7.0970441026343978E-5,-0.081048819235342642,-0.00024549134958053907,-1.7425575551665338E-5,0.0,0.0,0.0,0.0,0.0,0.0,
        0.0,0.0,0.093363604583182686,3.0799370827412689E-5,-0.00012782334615158236,-0.032334731686097067,
        -2.0477343242432103E-7,1.7896052771145248E-5,-0.024963107708841741,-1.6194155578034896E-5,0.00015880460924100231,
        -0.020118546073300689,-2.667646069196824E-5,0.0,0.0,0.0,0.0,0.0,0.0,0.0,0.0,0.0,0.49813926195152913,
        -0.00017528152484155724,0.00018393080016621108,-0.17188619370616637,-9.4178350536048286E-5,0.00017435004524606152,
        -0.13298344865537265,-1.2401466248264971E-5,0.00016997199450951656,-0.10796159984175095,0.0,0.0,0.0,0.0,0.0,0.0,0.0,
        0.0,0.0,0.0,0.39535959807028387,-0.00099043984756774762,-0.00016984196181567382,-0.10065418304586403,
        -0.001039333890452857,-0.00014846960874629052,-0.082085488838510676,-0.00088014262683248272,-0.00011298643072860384,
        0.0,0.0,0.0,0.0,0.0,0.0,0.0,0.0,0.0,0.0,0.0,0.098784373897778111,1.379925875586597E-5,-0.00021307203223217444,
        -0.025317508154544546,-3.8586189065682468E-6,-0.00010205938740070629,-0.020627333316023115,-1.5190280508914674E-5,0.0,
        0.0,0.0,0.0,0.0,0.0,0.0,0.0,0.0,0.0,0.0,0.0,0.52749981350157449,-0.00023432812992100008,0.00011672307002264918,
        -0.13343842177106774,-0.00016911926055907214,0.00013367833808069503,-0.10882333220692945,0.0,0.0,0.0,0.0,0.0,0.0,0.0,
        0.0,0.0,0.0,0.0,0.0,0.0,0.40767379600460241,-0.001420492715637155,-0.00022515367522466954,-0.083125610401955277,
        -0.0014882250041309344,-0.00020821798398764949,0.0,0.0,0.0,0.0,0.0,0.0,0.0,0.0,0.0,0.0,0.0,0.0,0.0,0.0,
        0.10177053391227749,8.63137591583232E-6,-0.0003630007358021759,-0.021130857297298654,-3.5781330140089059E-6,0.0,0.0,
        0.0,0.0,0.0,0.0,0.0,0.0,0.0,0.0,0.0,0.0,0.0,0.0,0.0,0.544082295885682,-0.000326621182822086,9.4506531633399324E-5,
        -0.10972642159828502,0.0,0.0,0.0,0.0,0.0,0.0,0.0,0.0,0.0,0.0,0.0,0.0,0.0,0.0,0.0,0.0,0.41538729066323726,
        -0.0020700877740851965,-0.00030221634851523653,0.0,0.0,0.0,0.0,0.0,0.0,0.0,0.0,0.0,0.0,0.0,0.0,0.0,0.0,0.0,0.0,0.0,
        0.10358194532626247,8.2420493374344387E-6,0.0,0.0,0.0,0.0,0.0,0.0,0.0,0.0,0.0,0.0,0.0,0.0,0.0,0.0,0.0,0.0,0.0,0.0,
        0.554556561972674,0.0,0.0,0.0,0.0,0.0,0.0,0.0,0.0,0.0,0.0,0.0,0.0,0.0,0.0,0.0,0.0,0.0,0.0,0.0,0.003162277660168379];
    MPC_3_f_a: ARRAY [0..20] OF REAL := [1.322628327144006E-6,-0.00048116811531683895,-4.3296165052708516E-6,-55.375904267141834,
        0.0,0.0,0.0,-6.9150559684644062E-11,3.7716284508284807E-8,-0.0027971712823564414,-78.996564422017926,0.0,0.0,0.0,
        -2.394037186466665E-10,1.3057639972340998E-7,2.8628831792336135E-7,-273.49234867499621,0.0,0.0,0.0];
    MPC_3_g_a: ARRAY [0..20] OF REAL := [-0.0812759988320282,0.12878974211545094,0.004723574350295019,1608.467976495617,
        3.4881337436777868,-1.3447885799979735,-1.1731438171326984,0.27540380820784305,0.004147779263663315,0.10291146104511424,
        371.46041919189759,0.11111867957141465,2.7949959088743945,-2.8155753844244238,0.065710282048828311,0.023308594370287667,
        0.00655318586773693,16000.578760709672,1.6106730948139927,2.3311020292522739,2.4089351935793255];
    MPC_3_e_a: ARRAY [0..48] OF REAL := [0.9945076508163887,-7.4955911032675407E-6,0.018219343923005435,-0.86686845021470726,0.0,
        0.0,0.0,-0.0054923962532121753,0.99999067551082088,0.018219326989996565,-1.077349693812959,0.0,0.0,0.0,
        -4.0627503649808205E-13,2.2159162199695515E-10,0.99998342284905262,-0.4641225044555104,0.0,0.0,0.0,2.6237854624951297E-12,
        -9.54430195553142E-10,-2.0954813586927272E-9,0.99929334159686478,0.0,0.0,0.0,-6.3159654022047717E-6,0.0022977287773259252,
        2.0675277771461239E-5,264.43732399282771,1.0,0.0,0.0,0.002815004563879495,-1.3684281447907272E-7,2.54613431540441E-5,264.43733847702208,
        0.0,1.0,0.0,2.3147841327022809E-10,-1.26253752403586E-7,-2.7681092818992033E-7,264.43856123334115,0.0,0.0,1.0];
    i0_mpcblock_refmd: mpcblock_refmd_MPC;
    i0_mpc_clipping: mpc_clipping_MPC;
    i0_qr: qr_MPC;
    i0_maximum2: maximum2_MPC;
    i0_DropConstraint: DropConstraint_MPC;
    i0_b_abs: b_abs_MPC;
    i0_abs_g: abs_g_MPC;
    xk: ARRAY [0..6] OF REAL;
    y_innov: ARRAY [0..2] OF REAL;
    v: REAL;
    rseq: ARRAY [0..2] OF REAL;
    aZZ1: ARRAY [0..71] OF REAL;
    zopt: ARRAY [0..18] OF REAL;
    b_i: DINT;
    b_b: ARRAY [0..71] OF REAL;
    b_r: ARRAY [0..18] OF REAL;
    rMin: REAL;
    b_H: ARRAY [0..360] OF REAL;
    cTol: ARRAY [0..71] OF REAL;
    cTolComputed: BOOL;
    iC: ARRAY [0..71] OF DINT;
    nA: DINT;
    Opt: ARRAY [0..37] OF REAL;
    Rhs: ARRAY [0..37] OF REAL;
    DualFeasible: BOOL;
    tmp: DINT;
    ColdReset: BOOL;
    kDrop: DINT;
    Xnorm0: REAL;
    cMin: REAL;
    cVal: REAL;
    z: ARRAY [0..18] OF REAL;
    t: REAL;
    iSave: DINT;
    w_i: DINT;
    j_k: DINT;
    rtb_iAout: ARRAY [0..71] OF BOOL;
    rtb_xest: ARRAY [0..6] OF REAL;
    b_Ac: ARRAY [0..18] OF REAL;
    old_u: ARRAY [0..2] OF REAL;
    iC_0: DINT;
    y_innov_0: REAL;
    b_H_tmp: DINT;
    D_tmp: DINT;
    exitg1: DINT;
    exitg2: DINT;
    exitg3: DINT;
    exitg4: DINT;
    temp1: BOOL;
    temp4: ARRAY [0..18] OF REAL;
    temp5: REAL;
    temp6: ARRAY [0..71] OF REAL;
END_VAR
VAR_TEMP
    (* Matrices de trabajo del QP: en cada ejecucion se escriben antes de leerse *)
    RLinv: ARRAY [0..360] OF REAL;
    TL: ARRAY [0..360] OF REAL;
    b_D: ARRAY [0..360] OF REAL;
END_VAR
CASE ssMethodType OF
    0:
        PLCGlobalVarMPC.plc_ts_counter_MPC := 0;
        (* SystemInitialize for Atomic SubSystem: '<Root>/MPC_3' *)
        (* InitializeConditions for Memory: '<S3>/Memory' *)
        FOR kDrop := 0 TO 71 DO
            Memory_PreviousInput[kDrop] := FALSE;
        END_FOR;
        (* End of InitializeConditions for Memory: '<S3>/Memory' *)

        (* InitializeConditions for UnitDelay: '<S3>/last_mv' *)
        last_mv_DSTATE[0] := 0.656128124791873;
        last_mv_DSTATE[1] := 0.23798560261559079;
        last_mv_DSTATE[2] := 0.47436402610926476;
        (* End of SystemInitialize for SubSystem: '<Root>/MPC_3' *)
        (* SystemInitialize for Atomic SubSystem: '<Root>/MPC_3' *)
        (* InitializeConditions for Memory: '<S3>/last_x' *)
        FOR kDrop := 0 TO 6 DO
            last_x_PreviousInput[kDrop] := c_last_x_InitialCond[kDrop];
        END_FOR;
        (* End of InitializeConditions for Memory: '<S3>/last_x' *)
        (* End of SystemInitialize for SubSystem: '<Root>/MPC_3' *)

        (* ConstCode for Atomic SubSystem: '<Root>/MPC_3' *)
        (* ConstCode for Math: '<S3>/Math Function' incorporates:
         *  Constant: '<S2>/y.wt_zero' *)
        MathFunction[0] := 0.0;
        (* ConstCode for Math: '<S3>/Math Function1' incorporates:
         *  Constant: '<S2>/u.wt_zero' *)
        MathFunction1[0] := 0.0;
        (* ConstCode for Math: '<S3>/Math Function2' incorporates:
         *  Constant: '<S2>/du.wt_zero' *)
        MathFunction2[0] := 0.0;
        (* ConstCode for Math: '<S3>/Math Function' incorporates:
         *  Constant: '<S2>/y.wt_zero' *)
        MathFunction[1] := 0.0;
        (* ConstCode for Math: '<S3>/Math Function1' incorporates:
         *  Constant: '<S2>/u.wt_zero' *)
        MathFunction1[1] := 0.0;
        (* ConstCode for Math: '<S3>/Math Function2' incorporates:
         *  Constant: '<S2>/du.wt_zero' *)
        MathFunction2[1] := 0.0;
        (* ConstCode for Math: '<S3>/Math Function' incorporates:
         *  Constant: '<S2>/y.wt_zero' *)
        MathFunction[2] := 0.0;
        (* ConstCode for Math: '<S3>/Math Function1' incorporates:
         *  Constant: '<S2>/u.wt_zero' *)
        MathFunction1[2] := 0.0;
        (* ConstCode for Math: '<S3>/Math Function2' incorporates:
         *  Constant: '<S2>/du.wt_zero' *)
        MathFunction2[2] := 0.0;
        (* End of ConstCode for SubSystem: '<Root>/MPC_3' *)
    1:
        IF PLCGlobalVarMPC.plc_ts_counter_MPC = 0 THEN
            (* [DIAG] inicio de la medicion *)
            "Diag_HIL".mpc_aux := RUNTIME("Diag_HIL".mpc_mem);

